// TIA Portal V20 export
// export: Created 2026-10-19T18:37:59.2059828Z, ExportSetting WithDefaults, DisplayName Totally Integrated Automation Portal, DisplayVersion V20 Update 6, DisplayName TIA Portal Openness, DisplayVersion V20 Update 6, DisplayName TIA Portal Version Control Interface, DisplayVersion V20 Update 6, DisplayName SINAMICS Startdrive Advanced, DisplayVersion V20 SP1, DisplayName SINAMICS Startdrive G130, G150, S120, S150, SINAMICS MV, G220, S200, S210, DisplayVersion V20 SP1, DisplayName SINAMICS Startdrive G110M, G120, G120C, G120D, G120P, G115D, DisplayVersion V20 SP1, DisplayName STEP 7 Professional, DisplayVersion V20 Update 6, DisplayName STEP 7 Safety, DisplayVersion V20 Update 2, DisplayName WinCC Basic/Comfort/Advanced, DisplayVersion V20 Update 6, DisplayName WinCC Unified, DisplayVersion V20 Update 6
DATA_BLOCK "Order_Table_Buffers_FB_DB_2"   // DB19
VERSION : 0.1
// stored: AutoNumber true, DBAccessibleFromOPCUA true, InstanceOfName Order_Table_Buffers_FB, InstanceOfType FB
"Order_Table_Buffers_FB"
   // VAR_INPUT
   //    System_Selected { ExternalWritable := 'False'} : Bool;
   //    AutoMan_Switch : Bool;
   //    CurrentTime { ExternalWritable := 'False'} : String;
   //    CurrentDTL : DTL;
   //    Watchdog : "Watchdog_Settings_UDT";
   //    VTD_CurrentLevel : UInt;
   //    OPC_UA_State_VTD : UInt;
   //    OPC_UA_State_Main : UInt;
   //    OPC_UA_State_L2 : UInt;
   //    OPC_UA_State_L3 : UInt;
   //    OPC_UA_State_L4 : UInt;
   //    OPC_UA_State_L5 : UInt;
   //    OPC_UA_State_L6 : UInt;
   //    Clear_OrderTable : Bool;
   // END_VAR
   // VAR_IN_OUT
   //    Cnv_Buffer_21 : "Buffer_Cnv_Control";
   //    Cnv_Buffer_31 : "Buffer_Cnv_Control";
   //    Cnv_Buffer_41 : "Buffer_Cnv_Control";
   //    Cnv_Buffer_51 : "Buffer_Cnv_Control";
   //    Cnv_Buffer_61 : "Buffer_Cnv_Control";
   //    Cnv_Buffer_22 : "Buffer_Cnv_Control";
   //    Cnv_Buffer_32 : "Buffer_Cnv_Control";
   //    Cnv_Buffer_42 : "Buffer_Cnv_Control";
   //    Cnv_Buffer_52 : "Buffer_Cnv_Control";
   //    Cnv_Buffer_62 : "Buffer_Cnv_Control";
   //    System : "System_UDT";
   //    Control_OPC_Ua : "WMS_OPC_UA";
   // END_VAR
   // VAR
   //    L2_CurrentOrder { ExternalWritable := 'False'} : UDInt;
   //    L3_CurrentOrder : UDInt;
   //    L4_CurrentOrder : UDInt;
   //    L5_CurrentOrder : UDInt;
   //    L6_CurrentOrder : UDInt;
   //    L2DoneRTrig : R_TRIG;
   //    L3DoneRTrig { S7_SetPoint := 'True'} : R_TRIG;
   //    L4DoneRTrig { S7_SetPoint := 'True'} : R_TRIG;
   //    L5DoneRTrig { S7_SetPoint := 'True'} : R_TRIG;
   //    L6DoneRTrig { S7_SetPoint := 'True'} : R_TRIG;
   //    PalletRefused_RTrig { ExternalWritable := 'False'} : R_TRIG;
   //    ErrorRTrig { ExternalWritable := 'False'} : R_TRIG;
   //    CancelRTrig { ExternalWritable := 'False'} : R_TRIG;
   //    PauseRTrig { ExternalWritable := 'False'} : R_TRIG;
   //    ResumeRTrig { ExternalWritable := 'False'} : R_TRIG;
   //    Clear_Store : R_TRIG;
   //    Clear_Retrieve : R_TRIG;
   //    Canceling : Bool;
   //    L2_WatchdogTimer : TON_TIME;
   //    L3_WatchdogTimer { S7_SetPoint := 'True'} : TON_TIME;
   //    L4_WatchdogTimer { S7_SetPoint := 'True'} : TON_TIME;
   //    L5_WatchdogTimer { S7_SetPoint := 'True'} : TON_TIME;
   //    L6_WatchdogTimer { S7_SetPoint := 'True'} : TON_TIME;
   //    L2_WatchdogStart : Bool;
   //    L3_WatchdogStart : Bool;
   //    L4_WatchdogStart : Bool;
   //    L5_WatchdogStart : Bool;
   //    L6_WatchdogStart : Bool;
   //    F_AutoMode { S7_SetPoint := 'True'} : F_TRIG;
   // END_VAR
BEGIN
END_DATA_BLOCK
